// TIA Portal V20 program export: 0 tag tables, 0 data types, 0 data blocks, 2 code blocks (in call order from the OBs), 0 instance data blocks

ORGANIZATION_BLOCK "Main"   // OB1, SCL, ProgramCycle
{ S7_Optimized_Access := 'TRUE' }
// stored: SetENOAutomatically false
   VAR_INPUT
      Initial_Call : Bool;   // Initial call of this OB
      Remanence : Bool;   // =True, if remanent data are available
   END_VAR
BEGIN

   // Arnes de prueba para FC_Escalado (bloques-de-funcion/fc-escalado/arnes-ob1.md).
   //
   // Las seis variables de test son REAL: la API de PLCSIM Advanced resuelve y escribe
   // simbolos REAL de forma nativa, mientras que el bloque recibe INT. El arnes hace la
   // conversion con REAL_TO_INT, que trunca hacia cero, y los valores de prueba se
   // mantienen dentro del rango INT.
   //
   // Mapa de tags (tabla Agent_Escalado):
   //   RawValue    entrada  valor crudo de la entrada analogica
   //   RawMin      entrada  raw del minimo de escala
   //   RawMax      entrada  raw del maximo de escala
   //   ScaleMin    entrada  valor de ingenieria del raw minimo
   //   ScaleMax    entrada  valor de ingenieria del raw maximo
   //   ScaledValue salida   valor escalado
   "FC_Escalado"(iValorCrudo := REAL_TO_INT("RawValue"),
                 iRawMin := REAL_TO_INT("RawMin"),
                 iRawMax := REAL_TO_INT("RawMax"),
                 rEscalaMin := "ScaleMin",
                 rEscalaMax := "ScaleMax",
                 rEscalado => "ScaledValue");
END_ORGANIZATION_BLOCK

FUNCTION "FC_Escalado" : Void   // FC1, SCL
{ S7_Optimized_Access := 'TRUE' }
// ==============================================================================
//  Escala un valor analogico crudo a unidades de ingenieria.
// 
//  Es la pieza mas universal de cualquier proyecto con entradas analogicas: la
//  conversion 0-27648 -> 0.0-10.0 bar se reescribe en cada maquina y cada vez
//  aparecen los mismos errores: division por cero, overflow al restar, y el
//  cambio de INT a REAL hecho en el orden equivocado.
// 
//  Aqui la resta se hace EN REAL, no en INT: con el rango completo de INT
//  (-32768..32767) restar en INT puede desbordar y el resultado es un valor
//  sin sentido. La division por cero se cubre aparte y devuelve el minimo de
//  escala, que es la unica respuesta sensata cuando no hay rango.
// 
//  NO satura: si el raw esta fuera del rango configurado, el resultado sale
//  fuera de escala. Si necesitas saturar, envuelve la llamada con MIN/MAX.
// 
//  Consulta README.md de este recurso para la interfaz, las limitaciones y la
//  prueba ejecutada.
// ==============================================================================
// stored: SetENOAutomatically false
   VAR_INPUT
      iValorCrudo : Int;   // Valor crudo de la entrada analogica
      iRawMin : Int;   // Raw que corresponde al minimo de escala
      iRawMax : Int;   // Raw que corresponde al maximo de escala
      rEscalaMin : Real;   // Valor de ingenieria del raw minimo
      rEscalaMax : Real;   // Valor de ingenieria del raw maximo
   END_VAR
   VAR_OUTPUT
      rEscalado : Real;   // Valor escalado en unidades de ingenieria
   END_VAR
BEGIN


   // Sin rango no hay escala posible: se devuelve el minimo en vez de dejar que
   // la division por cero reviente el ciclo.
   IF #iRawMax = #iRawMin THEN
       #rEscalado := #rEscalaMin;
   ELSE
       #rEscalado := #rEscalaMin
       + ((INT_TO_REAL(#iValorCrudo) - INT_TO_REAL(#iRawMin))
       / (INT_TO_REAL(#iRawMax) - INT_TO_REAL(#iRawMin)))
       * (#rEscalaMax - #rEscalaMin);
   END_IF;
END_FUNCTION
